(* IEC 61131-3 sources: plc-vscode/tests/st/all/trust-platform/examples/OSCAT/airport_baggage_command_observer/oop/src, 3 files *)

(* ---- Main.st ---- *)
(* Pattern role: IBaggageCommand is the contract boundary for the Command and Observer example. *)
INTERFACE IBaggageCommand
    PROPERTY CommandId : INT
    GET
    END_GET
    END_PROPERTY
    METHOD Execute : BOOL
    VAR_INPUT
        BagId : INT;
    END_VAR
    END_METHOD
END_INTERFACE

(* Pattern role: IBaggageEventSubscriber is the contract boundary for the Command and Observer example. *)
INTERFACE IBaggageEventSubscriber
    METHOD OnBaggageEvent
    VAR_INPUT
        BagId : INT;
        CommandId : INT;
    END_VAR
    END_METHOD
END_INTERFACE

(* Pattern role: DivertLeftCommand is a concrete implementation in the Command and Observer example. *)
FUNCTION_BLOCK DivertLeftCommand IMPLEMENTS IBaggageCommand
METHOD PUBLIC Execute : BOOL
VAR_INPUT
    BagId : INT;
END_VAR
Execute := TRUE;
END_METHOD
PUBLIC PROPERTY CommandId : INT
GET
    CommandId := INT#1;
END_GET
END_PROPERTY
END_FUNCTION_BLOCK

(* Pattern role: DivertRightCommand is a concrete implementation in the Command and Observer example. *)
FUNCTION_BLOCK DivertRightCommand IMPLEMENTS IBaggageCommand
METHOD PUBLIC Execute : BOOL
VAR_INPUT
    BagId : INT;
END_VAR
Execute := TRUE;
END_METHOD
PUBLIC PROPERTY CommandId : INT
GET
    CommandId := INT#2;
END_GET
END_PROPERTY
END_FUNCTION_BLOCK

(* Pattern role: RejectBagCommand is a concrete implementation in the Command and Observer example. *)
FUNCTION_BLOCK RejectBagCommand IMPLEMENTS IBaggageCommand
METHOD PUBLIC Execute : BOOL
VAR_INPUT
    BagId : INT;
END_VAR
Execute := TRUE;
END_METHOD
PUBLIC PROPERTY CommandId : INT
GET
    CommandId := INT#3;
END_GET
END_PROPERTY
END_FUNCTION_BLOCK

(* Pattern role: BaggageHistorianSubscriber is a concrete implementation in the Command and Observer example. *)
FUNCTION_BLOCK BaggageHistorianSubscriber IMPLEMENTS IBaggageEventSubscriber
VAR
    EventCountValue : INT;
END_VAR
METHOD PUBLIC OnBaggageEvent
VAR_INPUT
    BagId : INT;
    CommandId : INT;
END_VAR
EventCountValue := EventCountValue + INT#1;
END_METHOD
PUBLIC PROPERTY EventCount : INT
GET
    EventCount := EventCountValue;
END_GET
END_PROPERTY
END_FUNCTION_BLOCK

(* Pattern role: BaggageMqttSubscriber is a concrete implementation in the Command and Observer example. *)
FUNCTION_BLOCK BaggageMqttSubscriber IMPLEMENTS IBaggageEventSubscriber
VAR
    PublishReadyValue : BOOL;
END_VAR
METHOD PUBLIC OnBaggageEvent
VAR_INPUT
    BagId : INT;
    CommandId : INT;
END_VAR
PublishReadyValue := TRUE;
END_METHOD
PUBLIC PROPERTY PublishReady : BOOL
GET
    PublishReady := PublishReadyValue;
END_GET
END_PROPERTY
END_FUNCTION_BLOCK

(* Composition role: BaggageEventBus owns the collaborating objects used by this Command and Observer example. *)
FUNCTION_BLOCK BaggageEventBus
VAR
    Historian : IBaggageEventSubscriber;
    Mqtt : IBaggageEventSubscriber;
END_VAR
METHOD PUBLIC Subscribe
VAR_INPUT
    HistorianSub : IBaggageEventSubscriber;
    MqttSub : IBaggageEventSubscriber;
END_VAR
Historian := HistorianSub;
Mqtt := MqttSub;
END_METHOD
METHOD PUBLIC Publish
VAR_INPUT
    BagId : INT;
    CommandId : INT;
END_VAR
Historian.OnBaggageEvent(BagId := BagId, CommandId := CommandId);
Mqtt.OnBaggageEvent(BagId := BagId, CommandId := CommandId);
END_METHOD
END_FUNCTION_BLOCK

(* Composition role: BaggageDiverter owns the collaborating objects used by this Command and Observer example. *)
FUNCTION_BLOCK BaggageDiverter
VAR
    Left : DivertLeftCommand;
    Right : DivertRightCommand;
    Reject : RejectBagCommand;
    CurrentCommand : IBaggageCommand;
    Bus : BaggageEventBus;
    Historian : BaggageHistorianSubscriber;
    Mqtt : BaggageMqttSubscriber;
    LastBagIdValue : INT;
    LastCommandIdValue : INT;
END_VAR
METHOD PUBLIC Initialize
Bus.Subscribe(HistorianSub := Historian, MqttSub := Mqtt);
END_METHOD
METHOD PUBLIC SelectCommand : IBaggageCommand
VAR_INPUT
    ScannerResult : INT;
END_VAR
IF ScannerResult = INT#1 THEN
    SelectCommand := Left;
ELSIF ScannerResult = INT#2 THEN
    SelectCommand := Right;
ELSE
    SelectCommand := Reject;
END_IF;
END_METHOD
METHOD PUBLIC ProcessBag : INT
VAR_INPUT
    BagId : INT;
    ScannerResult : INT;
END_VAR
CurrentCommand := SelectCommand(ScannerResult := ScannerResult);
IF CurrentCommand.Execute(BagId := BagId) THEN
    LastBagIdValue := BagId;
    LastCommandIdValue := CurrentCommand.CommandId;
    Bus.Publish(BagId := BagId, CommandId := LastCommandIdValue);
END_IF;
ProcessBag := LastCommandIdValue;
END_METHOD
PUBLIC PROPERTY LastBagId : INT
GET
    LastBagId := LastBagIdValue;
END_GET
END_PROPERTY
PUBLIC PROPERTY LastCommandId : INT
GET
    LastCommandId := LastCommandIdValue;
END_GET
END_PROPERTY
PUBLIC PROPERTY EventCount : INT
GET
    EventCount := Historian.EventCount;
END_GET
END_PROPERTY
PUBLIC PROPERTY MqttPublishReady : BOOL
GET
    MqttPublishReady := Mqtt.PublishReady;
END_GET
END_PROPERTY
END_FUNCTION_BLOCK

(* Scan role: Main wires the example objects and exposes the PLC call path under test. *)
PROGRAM Main
VAR
    Diverter : BaggageDiverter;
    BagIdRaw : INT;
    ScannerResultRaw : INT;
    LeftOut : BOOL;
    RightOut : BOOL;
    RejectOut : BOOL;
END_VAR
Diverter.Initialize();
Diverter.ProcessBag(BagId := BagIdRaw, ScannerResult := ScannerResultRaw);
LeftOut := Diverter.LastCommandId = INT#1;
RightOut := Diverter.LastCommandId = INT#2;
RejectOut := Diverter.LastCommandId = INT#3;
END_PROGRAM

(* ---- Configuration.st ---- *)
CONFIGURATION AirportBaggageCommandObserverOopConfiguration
RESOURCE Cpu0 ON PLC
    TASK MainTask (INTERVAL := T#50ms, PRIORITY := 1);
    PROGRAM Diverter WITH MainTask : Main;
END_RESOURCE
VAR_CONFIG
    Diverter.BagIdRaw AT %IW0 : INT;
    Diverter.ScannerResultRaw AT %IW2 : INT;
    Diverter.LeftOut AT %QX0.0 : BOOL;
    Diverter.RightOut AT %QX0.1 : BOOL;
    Diverter.RejectOut AT %QX0.2 : BOOL;
END_VAR
END_CONFIGURATION

(* ---- Tests.st ---- *)
TEST_PROGRAM BaggageCommandExecutesScannerDecision
VAR
    Diverter : BaggageDiverter;
END_VAR
Diverter.Initialize();
ASSERT_EQUAL(EXPECTED := INT#2, ACTUAL := Diverter.ProcessBag(BagId := INT#42, ScannerResult := INT#2));
ASSERT_EQUAL(EXPECTED := INT#42, ACTUAL := Diverter.LastBagId);
END_TEST_PROGRAM

TEST_PROGRAM BaggageObserverPublishesAuditEvent
VAR
    Diverter : BaggageDiverter;
END_VAR
Diverter.Initialize();
Diverter.ProcessBag(BagId := INT#43, ScannerResult := INT#9);
ASSERT_EQUAL(EXPECTED := INT#1, ACTUAL := Diverter.EventCount);
ASSERT_TRUE(IN := Diverter.MqttPublishReady);
ASSERT_EQUAL(EXPECTED := INT#3, ACTUAL := Diverter.LastCommandId);
END_TEST_PROGRAM

(* Multi-event scan-loop test: drives the diverter through several
   different scanner results and verifies the historian counts every
   event and LastBagId/LastCommandId reflect the most recent decision.
   Catches bugs where command selection or event publication leaks
   state between scans. *)
TEST_PROGRAM BaggageDiverterAccumulatesEventsAcrossScans
VAR
    Diverter : BaggageDiverter;
    I : INT;
END_VAR

Diverter.Initialize();

Diverter.ProcessBag(BagId := INT#1, ScannerResult := INT#1);
ASSERT_EQUAL(EXPECTED := INT#1, ACTUAL := Diverter.LastCommandId);
ASSERT_EQUAL(EXPECTED := INT#1, ACTUAL := Diverter.LastBagId);

Diverter.ProcessBag(BagId := INT#2, ScannerResult := INT#2);
ASSERT_EQUAL(EXPECTED := INT#2, ACTUAL := Diverter.LastCommandId);
ASSERT_EQUAL(EXPECTED := INT#2, ACTUAL := Diverter.LastBagId);

Diverter.ProcessBag(BagId := INT#3, ScannerResult := INT#9);
ASSERT_EQUAL(EXPECTED := INT#3, ACTUAL := Diverter.LastCommandId);
ASSERT_EQUAL(EXPECTED := INT#3, ACTUAL := Diverter.LastBagId);

(* All three bags should have published to the historian *)
ASSERT_EQUAL(EXPECTED := INT#3, ACTUAL := Diverter.EventCount);
END_TEST_PROGRAM
